Fanuc KAREL source: ko00074.KL

-- PROVISIONAL review KL for V1013-1; original PC SHA256 df9d50bed4b2fdd0fc7b75dea68ca7211db50bd0ae633811afa66590a9f3dabe
-- Incomplete behavior may be omitted. Consult companion uncertainty JSON. Do not deploy.
PROGRAM KO00074
%NOLOCKGROUP
BEGIN
  -- UNRESOLVED_PC offsets 5-12; opcodes 9D,23
  -- UNRESOLVED_PC offsets 17-66; opcodes 27,22,1C,27,49,7E,AD,22,31,7E,4A
  -- UNRESOLVED_PC offsets 71-75; opcodes 7F
END KO00074
